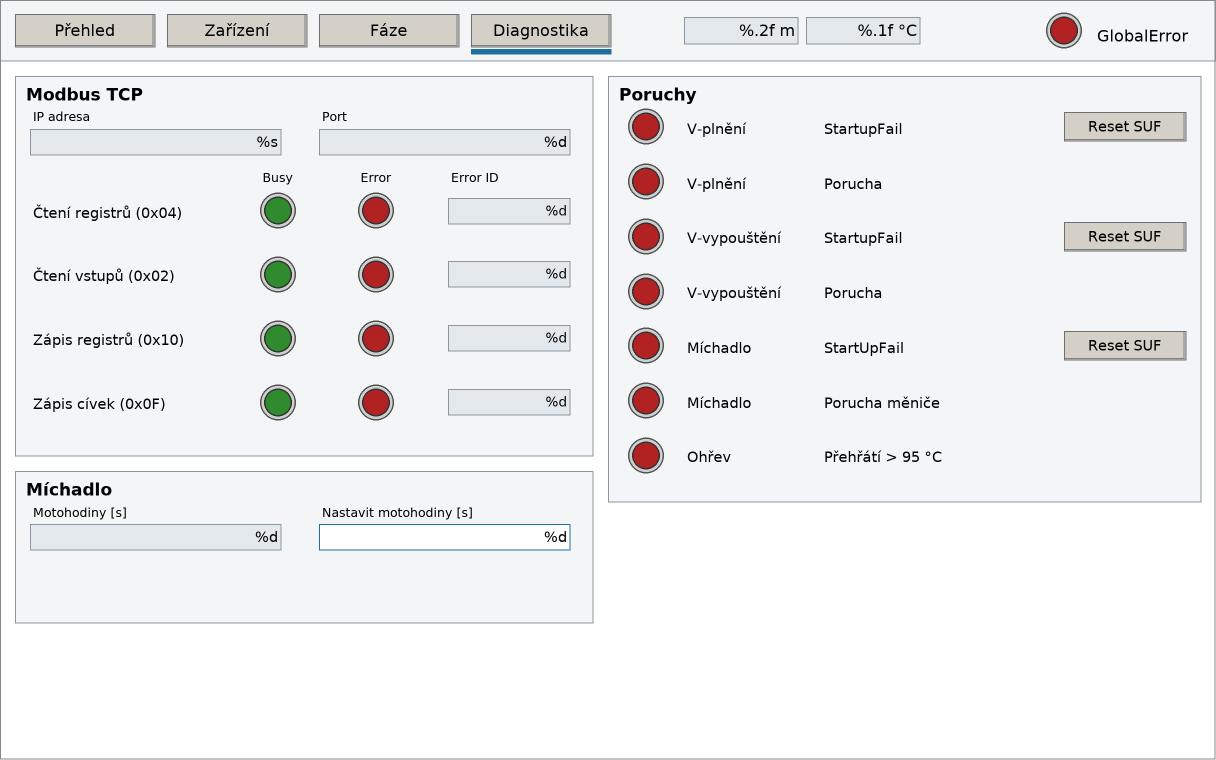
VISUALIZATION Diagnostika  // 1216x760
    Rectangle (0,0 1216x61)
    Button (15,14 140x33), "Přehled"
        OnMouseClick: change screen: Prehled
    Button (167,14 140x33), "Zařízení"
        OnMouseClick: change screen: Zarizeni
    Button (319,14 140x33), "Fáze"
        OnMouseClick: change screen: Faze
    Button (471,14 140x33), "Diagnostika"
        OnMouseClick: change screen: Diagnostika
    Rectangle (471,49 140x5)
    Rectangle (684,17 114x27), "%.2f m", text variable: Global.Tank1.Filling.WaterLevel
    Rectangle (806,17 114x27), "%.1f °C", text variable: Global.Tank1.Heating.WaterTemp
    Lamp1 (1041,10 46x41), variable: Global.Tank1.GlobalError, style: Lamp-Lamp1-Red
    Label (1094,23 126x26), "GlobalError"
    Rectangle (15,76 578x380)
    Label (23,81 122x27), "Modbus TCP"
    Label (30,106 83x21), "IP adresa"
    Rectangle (30,129 251x26), "%s", text variable: MB_Connector.mb_ipaddr
    Label (319,106 41x21), "Port"
    Rectangle (319,129 251x26), "%d", text variable: MB_Connector.mb_port
    Label (236,167 84x21), "Busy"
    Label (334,167 84x21), "Error"
    Label (433,167 84x21), "Error ID"
    Label (30,201 209x24), "Čtení registrů (0x04)"
    Lamp1 (255,190 46x41), variable: MB_Connector.mb_regs_busy, style: Lamp-Lamp1-Green
    Lamp1 (353,190 46x41), variable: MB_Connector.mb_regs_error, style: Lamp-Lamp1-Red
    Rectangle (448,198 122x26), "%d", text variable: MB_Connector.mb_regs_errid
    Label (30,264 190x24), "Čtení vstupů (0x02)"
    Lamp1 (255,254 46x41), variable: MB_Connector.mb_inps_busy, style: Lamp-Lamp1-Green
    Lamp1 (353,254 46x41), variable: MB_Connector.mb_inps_error, style: Lamp-Lamp1-Red
    Rectangle (448,261 122x26), "%d", text variable: MB_Connector.mb_inps_errid
    Label (30,328 209x24), "Zápis registrů (0x10)"
    Lamp1 (255,318 46x41), variable: MB_Connector.mbw_regs_busy, style: Lamp-Lamp1-Green
    Lamp1 (353,318 46x41), variable: MB_Connector.mbw_regs_error, style: Lamp-Lamp1-Red
    Rectangle (448,325 122x26), "%d", text variable: MB_Connector.mbw_regs_errid
    Label (30,392 180x24), "Zápis cívek (0x0F)"
    Lamp1 (255,382 46x41), variable: MB_Connector.mbw_coils_busy, style: Lamp-Lamp1-Green
    Lamp1 (353,382 46x41), variable: MB_Connector.mbw_coils_error, style: Lamp-Lamp1-Red
    Rectangle (448,389 122x26), "%d", text variable: MB_Connector.mbw_coils_errid
    Rectangle (608,76 593x426)
    Label (616,81 87x27), "Poruchy"
    Lamp1 (623,106 46x41), variable: Global.Tank1.ValveFilling.State.StartupFail, style: Lamp-Lamp1-Red
    Label (684,117 84x24), "V-plnění"
    Label (821,117 113x24), "StartupFail"
    Button (1064,112 122x29), "Reset SUF", colour toggle: Global.Tank1.ValveFilling.State.StartupFail
        tap Global.Tank1.ValveFilling.Cmd.ResetSUF
    Lamp1 (623,161 46x41), variable: Global.Tank1.ValveFilling.State.Err, style: Lamp-Lamp1-Red
    Label (684,172 84x24), "V-plnění"
    Label (821,172 74x24), "Porucha"
    Lamp1 (623,216 46x41), variable: Global.Tank1.ValveDraining.State.StartupFail, style: Lamp-Lamp1-Red
    Label (684,226 123x24), "V-vypouštění"
    Label (821,226 113x24), "StartupFail"
    Button (1064,222 122x29), "Reset SUF", colour toggle: Global.Tank1.ValveDraining.State.StartupFail
        tap Global.Tank1.ValveDraining.Cmd.ResetSUF
    Lamp1 (623,271 46x41), variable: Global.Tank1.ValveDraining.State.Err, style: Lamp-Lamp1-Red
    Label (684,281 123x24), "V-vypouštění"
    Label (821,281 74x24), "Porucha"
    Lamp1 (623,325 46x41), variable: Global.Tank1.Mixer.State.StartUpFail, style: Lamp-Lamp1-Red
    Label (684,336 84x24), "Míchadlo"
    Label (821,336 113x24), "StartUpFail"
    Button (1064,331 122x29), "Reset SUF", colour toggle: Global.Tank1.Mixer.State.StartUpFail
        tap Global.Tank1.Mixer.Cmd.ResetSUF
    Lamp1 (623,380 46x41), variable: Global.Tank1.Mixer.State.Err, style: Lamp-Lamp1-Red
    Label (684,391 84x24), "Míchadlo"
    Label (821,391 142x24), "Porucha měniče"
    Lamp1 (623,435 46x41), variable: Global.Tank1.Heater.State.GenErr, style: Lamp-Lamp1-Red
    Label (684,445 55x24), "Ohřev"
    Label (821,445 161x24), "Přehřátí > 95 °C"
    Rectangle (15,471 578x152)
    Label (23,476 99x27), "Míchadlo"
    Label (30,502 125x21), "Motohodiny [s]"
    Rectangle (30,524 251x26), "%d", text variable: Global.Tank1.Mixer.State.RT
    Label (319,502 201x21), "Nastavit motohodiny [s]"
    Rectangle (319,524 251x26), "%d", text variable: Global.Tank1.Mixer.Cmd.SetRT
        OnMouseClick: write the text variable via Default
END_VISUALIZATION

(* stored: Version 1.1.0.1, ProductVersion 3.1.4024.16
   Visu Diagnostika: Id {07d02cde-6666-4b17-bfa0-f5de1ddc99be} *)
